(* IEC 61131-3 sources: st2fb/corpus_hard/unsupported_st/u05_pump_duty_records, 2 files *)

(* ---- control_flat.st ---- *)
(* Solvability control, never shown to a model: the same behaviour in the translator's v1 subset. Records became
   variables, EXIT became a loop condition. *)
FUNCTION_BLOCK PUMP_DUTY_SELECT
VAR_INPUT
  DEMAND : INT;
  AVAIL_1, AVAIL_2, AVAIL_3 : BOOL;
  RESET_TICKS : BOOL;
END_VAR
VAR_OUTPUT
  RUN_1, RUN_2, RUN_3 : BOOL;
  TICKS_1, TICKS_2, TICKS_3 : DINT;
  STARTS_TOTAL : INT;
  UNMET : INT;
END_VAR
VAR
  STARTS_1, STARTS_2, STARTS_3 : INT;
  WAS_1, WAS_2, WAS_3 : BOOL;
  PREV_DEMAND : INT;
  N : INT;
  BEST : INT;
  BEST_SCORE : DINT;
  SCORE : DINT;
  CHANGED : BOOL;
  SEARCHING : BOOL;
END_VAR
  CHANGED := (DEMAND <> PREV_DEMAND) OR (RUN_1 AND NOT AVAIL_1) OR (RUN_2 AND NOT AVAIL_2) OR (RUN_3 AND NOT AVAIL_3);
  PREV_DEMAND := DEMAND;

  IF CHANGED THEN
    WAS_1 := RUN_1;
    WAS_2 := RUN_2;
    WAS_3 := RUN_3;
    RUN_1 := FALSE;
    RUN_2 := FALSE;
    RUN_3 := FALSE;
    UNMET := 0;
    N := 1;
    SEARCHING := N <= DEMAND;
    WHILE SEARCHING DO
      BEST := 0;
      BEST_SCORE := 2147483647;
      IF AVAIL_1 AND NOT RUN_1 THEN
        SCORE := TICKS_1 + 5 * INT_TO_DINT(STARTS_1);
        IF SCORE < BEST_SCORE THEN
          BEST := 1;
          BEST_SCORE := SCORE;
        END_IF;
      END_IF;
      IF AVAIL_2 AND NOT RUN_2 THEN
        SCORE := TICKS_2 + 5 * INT_TO_DINT(STARTS_2);
        IF SCORE < BEST_SCORE THEN
          BEST := 2;
          BEST_SCORE := SCORE;
        END_IF;
      END_IF;
      IF AVAIL_3 AND NOT RUN_3 THEN
        SCORE := TICKS_3 + 5 * INT_TO_DINT(STARTS_3);
        IF SCORE < BEST_SCORE THEN
          BEST := 3;
          BEST_SCORE := SCORE;
        END_IF;
      END_IF;
      CASE BEST OF
        0:
          UNMET := DEMAND - N + 1;
          SEARCHING := FALSE;
        1:
          RUN_1 := TRUE;
          IF NOT WAS_1 THEN
            STARTS_1 := STARTS_1 + 1;
            STARTS_TOTAL := STARTS_TOTAL + 1;
          END_IF;
        2:
          RUN_2 := TRUE;
          IF NOT WAS_2 THEN
            STARTS_2 := STARTS_2 + 1;
            STARTS_TOTAL := STARTS_TOTAL + 1;
          END_IF;
        3:
          RUN_3 := TRUE;
          IF NOT WAS_3 THEN
            STARTS_3 := STARTS_3 + 1;
            STARTS_TOTAL := STARTS_TOTAL + 1;
          END_IF;
      END_CASE;
      N := N + 1;
      IF N > DEMAND THEN
        SEARCHING := FALSE;
      END_IF;
    END_WHILE;
  END_IF;

  IF RESET_TICKS THEN
    TICKS_1 := 0;
    TICKS_2 := 0;
    TICKS_3 := 0;
  ELSE
    IF RUN_1 THEN
      TICKS_1 := TICKS_1 + 1;
    END_IF;
    IF RUN_2 THEN
      TICKS_2 := TICKS_2 + 1;
    END_IF;
    IF RUN_3 THEN
      TICKS_3 := TICKS_3 + 1;
    END_IF;
  END_IF;
END_FUNCTION_BLOCK

(* ---- program.st ---- *)
(* Duty selection over pump records. *)
TYPE
  PUMP_RECORD : STRUCT
    AVAILABLE : BOOL;
    RUNNING : BOOL;
    RUN_TICKS : DINT;
    STARTS : INT;
  END_STRUCT;
END_TYPE

FUNCTION_BLOCK PUMP_DUTY_SELECT
VAR_INPUT
  DEMAND : INT;
  AVAIL_1, AVAIL_2, AVAIL_3 : BOOL;
  RESET_TICKS : BOOL;
END_VAR
VAR_OUTPUT
  RUN_1, RUN_2, RUN_3 : BOOL;
  TICKS_1, TICKS_2, TICKS_3 : DINT;
  STARTS_TOTAL : INT;
  UNMET : INT;
END_VAR
VAR CONSTANT
  PUMP_COUNT : INT := 3;
  WEAR_PER_START : DINT := 5;
END_VAR
VAR
  PUMP : ARRAY[1..3] OF PUMP_RECORD;
  PREV_DEMAND : INT;
  N, P : INT;
  WAS_RUNNING : ARRAY[1..3] OF BOOL;
END_VAR
VAR_TEMP
  BEST : INT;
  BEST_SCORE : DINT;
  SCORE : DINT;
  CHANGED : BOOL;
END_VAR
  PUMP[1].AVAILABLE := AVAIL_1;
  PUMP[2].AVAILABLE := AVAIL_2;
  PUMP[3].AVAILABLE := AVAIL_3;

  (* Reselect when demand changes, or when a running pump has become unavailable. *)
  CHANGED := DEMAND <> PREV_DEMAND;
  FOR P := 1 TO PUMP_COUNT DO
    IF PUMP[P].RUNNING AND NOT PUMP[P].AVAILABLE THEN
      CHANGED := TRUE;
      EXIT;
    END_IF;
  END_FOR;
  PREV_DEMAND := DEMAND;

  IF CHANGED THEN
    FOR P := 1 TO PUMP_COUNT DO
      WAS_RUNNING[P] := PUMP[P].RUNNING;
      PUMP[P].RUNNING := FALSE;
    END_FOR;
    UNMET := 0;
    FOR N := 1 TO DEMAND DO
      BEST := 0;
      BEST_SCORE := 2147483647;
      FOR P := 1 TO PUMP_COUNT DO
        IF PUMP[P].AVAILABLE AND NOT PUMP[P].RUNNING THEN
          SCORE := PUMP[P].RUN_TICKS + WEAR_PER_START * INT_TO_DINT(PUMP[P].STARTS);
          IF SCORE < BEST_SCORE THEN
            BEST := P;
            BEST_SCORE := SCORE;
          END_IF;
        END_IF;
      END_FOR;
      IF BEST = 0 THEN
        UNMET := DEMAND - N + 1;
        EXIT;
      END_IF;
      PUMP[BEST].RUNNING := TRUE;
      IF NOT WAS_RUNNING[BEST] THEN
        PUMP[BEST].STARTS := PUMP[BEST].STARTS + 1;
        STARTS_TOTAL := STARTS_TOTAL + 1;
      END_IF;
    END_FOR;
  END_IF;

  FOR P := 1 TO PUMP_COUNT DO
    IF RESET_TICKS THEN
      PUMP[P].RUN_TICKS := 0;
    ELSIF PUMP[P].RUNNING THEN
      PUMP[P].RUN_TICKS := PUMP[P].RUN_TICKS + 1;
    END_IF;
  END_FOR;

  RUN_1 := PUMP[1].RUNNING;
  RUN_2 := PUMP[2].RUNNING;
  RUN_3 := PUMP[3].RUNNING;
  TICKS_1 := PUMP[1].RUN_TICKS;
  TICKS_2 := PUMP[2].RUN_TICKS;
  TICKS_3 := PUMP[3].RUN_TICKS;
END_FUNCTION_BLOCK
